(* IEC 61131-3 sources: llm-plc-st-eval/data/processed_definitivo/gpt-4o-2024-08-06/B3/zero_shot, 3 files *)

(* ---- ejec_1.st ---- *)
FUNCTION_BLOCK FB_Contador
VAR_INPUT
    sensorPieza : BOOL;   // Entrada del sensor fotoeléctrico
    btnReset : BOOL;      // Botón de reset
END_VAR

VAR_OUTPUT
    loteListo : BOOL;     // Salida que indica si el lote está completo
    cuenta : INT;         // Contador de piezas
END_VAR

VAR
    sensorPiezaAnt : BOOL; // Estado anterior del sensor
END_VAR

// Inicialización de variables
sensorPiezaAnt := FALSE;
cuenta := 0;
loteListo := FALSE;

// Cuerpo del bloque de función
IF btnReset THEN
    // Si se presiona el botón de reset, reiniciar el contador y la salida de lote
    cuenta := 0;
    loteListo := FALSE;
ELSE
    // Detectar flanco ascendente del sensor
    IF (sensorPieza AND NOT sensorPiezaAnt) THEN
        // Incrementar el contador al detectar una pieza
        cuenta := cuenta + 1;
    END_IF;

    // Verificar si se ha completado el lote
    IF cuenta >= 12 THEN
        loteListo := TRUE;
    ELSE
        loteListo := FALSE;
    END_IF;
END_IF;

// Actualizar el estado anterior del sensor
sensorPiezaAnt := sensorPieza;

END_FUNCTION_BLOCK

(* ---- ejec_2.st ---- *)
FUNCTION_BLOCK FB_Contador
VAR_INPUT
    sensorPieza : BOOL;   // Entrada del sensor fotoeléctrico
    btnReset : BOOL;      // Botón de reset
END_VAR

VAR_OUTPUT
    loteListo : BOOL;     // Indica si el lote está completo
    cuenta : INT;         // Cuenta de piezas detectadas
END_VAR

VAR
    prevSensorPieza : BOOL; // Estado previo del sensor
END_VAR

// Inicialización de variables
IF btnReset THEN
    cuenta := 0;          // Reinicia la cuenta si se presiona el botón de reset
    loteListo := FALSE;   // Desactiva la salida de lote completo
END_IF

// Detección de flanco ascendente del sensor
IF (NOT prevSensorPieza) AND sensorPieza THEN
    cuenta := cuenta + 1; // Incrementa la cuenta al detectar una pieza
END_IF

// Comprobación de lote completo
IF cuenta >= 12 THEN
    loteListo := TRUE;    // Activa la salida de lote completo si se alcanzan 12 piezas
ELSE
    loteListo := FALSE;   // Asegura que la salida esté desactivada si no se alcanza el lote
END_IF

// Actualización del estado previo del sensor
prevSensorPieza := sensorPieza;

END_FUNCTION_BLOCK

(* ---- ejec_3.st ---- *)
FUNCTION_BLOCK FB_Contador
VAR_INPUT
    sensorPieza : BOOL;   // Entrada del sensor fotoeléctrico
    btnReset : BOOL;      // Botón de reset
END_VAR

VAR_OUTPUT
    loteListo : BOOL;     // Indica si el lote está completo
    cuenta : INT;         // Cuenta de piezas
END_VAR

VAR
    lastSensorState : BOOL; // Estado anterior del sensor
END_VAR

// Inicialización de variables
IF btnReset THEN
    cuenta := 0;
    loteListo := FALSE;
END_IF

// Detección de flanco ascendente del sensor
IF (sensorPieza AND NOT lastSensorState) THEN
    cuenta := cuenta + 1;
END_IF

// Comprobación si el lote está completo
IF cuenta >= 12 THEN
    loteListo := TRUE;
ELSE
    loteListo := FALSE;
END_IF

// Actualización del estado anterior del sensor
lastSensorState := sensorPieza;

END_FUNCTION_BLOCK
